(*
SPDX-FileCopyrightText: © 2026 Oleksandr Tiutyk <trofimich@gmail.com>
SPDX-License-Identifier: MIT
License: https://opensource.org/license/mit
*)

(*!
<summary>Checks interface-to-instance address conversion for a static object and for null.</summary>
<description>
Uses an owned static fixture. The converted address is borrowed and compared only in the calling task.
</description>
*)

{attribute 'no_assign'}
{attribute 'no_explicit_call' := 'do not call this function block directly'}
FUNCTION_BLOCK ObjectInterfaceAddressTest EXTENDS TOF_Testing.SingleCycleTest
VAR_STAT
	{attribute 'hide'}
	_ClassName : STRING := __POUNAME();
END_VAR
VAR
	_Probe : ObjectExitProbe;
END_VAR

(*!
<summary>Converts the live static interface, then checks that a null input does not reuse the address.</summary>
*)
METHOD PROTECTED ExecuteTest
VAR
	instance : TOF_Core.IObject;
END_VAR
instance := _Probe;
Assert.ThatBool(
	actual := TOF_Core.Memory.GetAddressFromInterface(interfaceInstance := instance) = ADR(_Probe),
	message := "The static interface must resolve to the complete probe address"
).IsTrue();

instance := 0;
Assert.ThatBool(
	actual := TOF_Core.Memory.GetAddressFromInterface(interfaceInstance := instance) = 0,
	message := "A null interface must return zero after a successful conversion"
).IsTrue();
END_METHOD

//! <summary>Borrows the concrete class name. Callers must not modify it.</summary>
{attribute 'monitoring' := 'call'}
PROPERTY ClassName : REFERENCE TO STRING
GET
ClassName REF= _ClassName;
END_GET
END_PROPERTY

//! <summary>Borrows the compiler-initialized namespace name. Callers must not modify it.</summary>
{attribute 'monitoring' := 'call'}
PROPERTY NamespaceName : REFERENCE TO STRING
GET
NamespaceName REF= CurrentNamespace.Name;
END_GET
END_PROPERTY

//! <summary>Reports the concrete instance size in bytes.</summary>
{attribute 'monitoring' := 'call'}
PROPERTY SelfSize : ULINT
GET
SelfSize := XSIZEOF(THIS^);
END_GET
END_PROPERTY

END_FUNCTION_BLOCK

(* stored: Version 1.1.0.1
   POU ObjectInterfaceAddressTest: Id {50301169-c256-4097-9740-c6af70175781}, SpecialFunc None
   Method ExecuteTest: Id {c3f58b6e-6421-4dd3-9590-a3d5650d5f05}
   Property ClassName: Id {65deeded-bb32-4287-beeb-73aebbde8ba9}
   Get Get: Id {7fc96a06-9ab4-4dd9-a0b1-1a76d7996a28}
   Property NamespaceName: Id {fb7385d6-619b-4c96-b677-967eaadb0aba}
   Get Get: Id {2a904551-d8a7-47b0-8c42-9690217eadcb}
   Property SelfSize: Id {5994c79d-bb34-4a5e-98c8-6dfd0a2f1a25}
   Get Get: Id {9612ca37-d224-40a4-8494-31cfefa1f0e2} *)
